(* IEC 61131-3 sources: esbmc-plc-benchmark-suite/benchmarks/manufacturing/st_counter_reset, 1 file *)

(* ---- counter_reset.st ---- *)
(* counter_reset: a free-running counter with a reset-to-value.
   Reset loads ResetCounterValue, otherwise Cnt increments; OUT follows Cnt.
   Imported from the Beremiz IEC 61131-3 language test (CounterST function block),
   re-expressed as a PROGRAM so it stands alone. See benchmark.yml for provenance. *)
PROGRAM drive
  VAR_INPUT
    Reset : BOOL;
    ResetCounterValue : INT;
  END_VAR
  VAR_OUTPUT
    OUT : INT;
  END_VAR
  VAR
    Cnt : INT;
  END_VAR

  IF Reset THEN
    Cnt := ResetCounterValue;
  ELSE
    Cnt := Cnt + 1;
  END_IF;

  OUT := Cnt;
END_PROGRAM
